// TIA Portal V21 program export: 0 tag tables, 0 data types, 0 data blocks, 2 code blocks (in call order from the OBs), 1 instance data blocks

ORGANIZATION_BLOCK "OB_Main"   // OB1, SCL, ProgramCycle
TITLE = "Main Program Sweep (Cycle)" / Main program of PLC_1200
{ S7_Optimized_Access := 'TRUE' }
// Calls the conveyor with the onboard inputs and output of the CPU 1214C
// stored: CodeModifiedDate 2026-10-23T19:59:16.3446293Z, CompileDate 2026-10-23T19:59:16.3446293Z, ConstantName OB_OB_Main, CreationDate 2026-10-23T19:59:09.2129607Z, DownloadDate 0001-01-01T00:00:00Z, EventClass Program cycle, InterfaceModifiedDate 2008-07-21T16:55:08.419547Z, IsConsistent true, LoadMemoryLength 4275, ModifiedDate 2026-10-23T19:59:16.3446293Z, ParameterModified 2008-07-21T16:55:08.419547Z, PriorityNumber 1, ProcessImagePartNumber 65535, SetENOAutomatically false, StructureModified 2008-07-21T16:55:08.419547Z, WorkMemoryLength 88
   VAR_INPUT
      Initial_Call : Bool;   // Initial call of this OB
      Remanence : Bool;   // =True, if remanent data are available
   END_VAR
BEGIN

       REGION Conveyor
           "IDB_Conveyor1200"(Start := "BeltStart",
                              Stop := "BeltStop",
                              SpeedRaw := "BeltSpeedRaw",
                              Motor => "BeltMotor");
       END_REGION
END_ORGANIZATION_BLOCK

FUNCTION_BLOCK "FB_Conveyor1200"   // FB1, SCL
TITLE = Conveyor on S7-1200
{ S7_Optimized_Access := 'TRUE' }
VERSION : 0.1
// TON exists on S7-1200 and S7-1500 alike. S7-1200 has no 64-bit data types (no LTime, LInt, LWord), so Time and DInt are used. SpeedRaw comes from the onboard analog input at %IW64 (0..27648).
// stored: AutoNumber true, IsIECCheckEnabled false, IsRetainMemResEnabled false, MemoryReserve 100, SetENOAutomatically false, UDAEnableTagReadback false
   VAR_INPUT
      Start : Bool;   // Start the belt
      Stop : Bool;   // Stop the belt
      SpeedRaw : Int;   // Raw value of the onboard analog input, 0..27648
   END_VAR
   VAR_OUTPUT
      Motor : Bool;   // Belt motor on
      Speed : Real;   // Belt speed in m/min
      DelayMilliseconds : DInt;   // Elapsed start delay in ms (DInt, no LInt on S7-1200)
   END_VAR
   VAR
      StartDelay { S7_SetPoint := 'True'} : TON_TIME;   // Start delay; TON_TIME, not TON_LTIME
      Running : Bool;   // Belt is commanded on
   END_VAR
   VAR CONSTANT
      RAW_FULL_SCALE : Int := 27648;   // Nominal range of the onboard analog input
      MAXIMUM_SPEED : Real := 30.0;   // Belt speed at full scale in m/min
   END_VAR
BEGIN

       REGION Command
           IF #Stop THEN
               #Running := FALSE;
           ELSIF #Start THEN
               #Running := TRUE;
           END_IF;
       END_REGION

       REGION Start delay and speed
           #StartDelay(IN := #Running, PT := T#2s);
           #Motor := #StartDelay.Q;
           #Speed := SCALE_X(MIN := 0.0, VALUE := NORM_X(MIN := 0, VALUE := #SpeedRaw, MAX := #RAW_FULL_SCALE), MAX := #MAXIMUM_SPEED);
           #DelayMilliseconds := TIME_TO_DINT(#StartDelay.ET);
       END_REGION
END_FUNCTION_BLOCK

DATA_BLOCK "IDB_Conveyor1200"   // DB1
VERSION : 0.1
// stored: AutoNumber true, DBAccessibleFromOPCUA true, InstanceOfName FB_Conveyor1200, InstanceOfType FB
"FB_Conveyor1200"
BEGIN
END_DATA_BLOCK
